{region 'Documentation'}
(*!
<summary>Owner execution and result snapshot.</summary>
*)
{endregion}
TYPE ST_ExecutionStatus :
STRUCT
    {attribute 'OPC.UA.DA.Access' := '1'}
    State : E_State := E_State.Uninitialized; //! Owner's detailed lifecycle state, including configured Test Case phases.
    {attribute 'OPC.UA.DA.Access' := '1'}
    ExecutionStatus : E_ExecutionStatus := E_ExecutionStatus.Unknown; //! Coarse execution classification derived from State.
    {attribute 'OPC.UA.DA.Access' := '1'}
    Result : E_Result := E_Result.NotEvaluated; //! Current held evaluation result; numeric order is not severity order.
    {attribute 'OPC.UA.DA.Access' := '1'}
    Uninitialized : BOOL := FALSE; //! Owner has not reached a reset-defined executable base state.
    {attribute 'OPC.UA.DA.Access' := '1'}
    ConfigError : BOOL := FALSE; //! Owner setup is invalid or has not yet been validated.
    {attribute 'OPC.UA.DA.Access' := '1'}
    Ready : BOOL := FALSE; //! Owner is initialized, Idle and ready to accept Start.
    {attribute 'OPC.UA.DA.Access' := '1'}
    Running : BOOL := FALSE; //! Owner is in its active execution phase.
    {attribute 'OPC.UA.DA.Access' := '1'}
    Completed : BOOL := FALSE; //! Owner has reached its terminal Completed state; does not imply Passed.
    {attribute 'OPC.UA.DA.Access' := '1'}
    Aborted : BOOL := FALSE; //! Owner completed with Abort result.
    {attribute 'OPC.UA.DA.Access' := '1'}
    // SA0033: Contract status field retained even when not consumed by this application.
    {attribute 'analysis' := '-33'}
    Inactive : BOOL := FALSE; //! Contract-reserved inactive indication; retained for compatible consumers.
    {attribute 'OPC.UA.DA.Access' := '1'}
    Error : BOOL := FALSE; //! Owner reports an error, including Result = Error.
END_STRUCT
END_TYPE

(* stored: Version 1.1.0.1
   DUT ST_ExecutionStatus: Id {731f2c13-6b9e-4d59-ab50-c6cf72fd3a3f} *)
